FUNCTION_BLOCK "FB_QualityEngine"
{ S7_Optimized_Access := 'TRUE' }
VERSION : 0.1

// Starter interface only. Confirm sensor scaling, target weights and sequence
// in TIA Portal and Machine Simulator before implementing quality decisions.

BEGIN
END_FUNCTION_BLOCK
